(* IEC 61131-3 sources: plc-st-coding-agent/progress/evidence/f14_v10_full_20261113/jobs/custom_minimax-m27 (part 3) *)

(* ---- public-hard-05.raw_candidate_01.st ---- *)
(* CONTRACT_RULES [] *)
FUNCTION_BLOCK ArmController
VAR_INPUT
    ManualMode      : BOOL;
    SingleStepMode  : BOOL;
    SingleCycleMode : BOOL;
    ContinuousMode  : BOOL;
    EmergencyStop   : BOOL;
    Start           : BOOL;
    DownButton      : BOOL;
    UpButton        : BOOL;
    LeftButton      : BOOL;
    RightButton     : BOOL;
    GripButton      : BOOL;
    ReleaseButton   : BOOL;
    DownLimitSwitch : BOOL;
    UpLimitSwitch   : BOOL;
    LeftLimitSwitch : BOOL;
    RightLimitSwitch: BOOL;
    GripLimitSwitch : BOOL;
    ReleaseLimitSwitch: BOOL;
END_VAR
VAR_OUTPUT
    MoveDown        : BOOL;
    MoveUp          : BOOL;
    MoveLeft        : BOOL;
    MoveRight       : BOOL;
    ActivateGrip    : BOOL;
    ActivateRelease : BOOL;
END_VAR
VAR
    tmp_Step : INT := 0;
    tmp_StartPrev : BOOL := FALSE;
    tmp_StartRisingEdge : BOOL;
    tmp_StartReleased : BOOL := FALSE;
    tmp_ActionCompleted : BOOL := FALSE;
END_VAR

(*
ENGINEERING_CONTRACT
====================================================================================================
Output State: Activation | Retention/hold | Explicit reset | Same-scan priority | Units/boundaries
----------------------------------------------------------------------------------------------------
MoveDown:     Manual=button AND NOT limit; Step modes=per step CASE; EmergencyStop→FALSE
MoveUp:       Manual=button AND NOT limit; Step modes=per step CASE; EmergencyStop→FALSE
MoveLeft:     Manual=button AND NOT limit; Step modes=per step CASE; EmergencyStop→FALSE
MoveRight:    Manual=button AND NOT limit; Step modes=per step CASE; EmergencyStop→FALSE
ActivateGrip:     Manual=GripButton; Step modes=per step CASE using GripLimitSwitch; EmergencyStop→FALSE
ActivateRelease:  Manual=ReleaseButton; Step modes=per step CASE using ReleaseLimitSwitch; EmergencyStop→FALSE

Manual Mode (PUB001):
  - Direct button-to-output mapping, held while button pressed and NOT at limit position
  - Grip/Release: held while button pressed (limit switches are feedback only)
  - Priority: Highest; independent of step sequencer state

Single Step Mode (PUB003):
  - Step sequence: Down→Grip→Up→Right→Down→Release→Up→Left→(repeat)
  - Each action requires limit switch confirmation before next Start enables next step
  - Initial arm position: top-left (UpLimitSwitch=1, LeftLimitSwitch=1) [PUB002]
  - Step 0: Wait for Start rising edge, then execute step 1
  - Steps 1-7: Advance when current action completes AND (Start released since last press OR step>0)
  - Step 8: Wait for Start released then pressed again before cycling to step 0

Single Cycle Mode (PUB005):
  - Auto-execute all 8 steps sequentially on single Start press
  - Stops at step 8 (end state) after completing left movement
  - No automatic restart; next Start press required

Continuous Mode (PUB006):
  - Same 8-step sequence as single cycle
  - Automatic restart from step 0 when left movement completes (step→0)
  - Continuous looping until mode change or emergency stop

Emergency Stop (PUB007):
  - Trigger: EmergencyStop=FALSE
  - Effect: All outputs FALSE, step counter reset to 0
  - No automatic resume; requires mode re-activation after E-stop clears

PUB IDs: PUB001, PUB002, PUB003, PUB004, PUB005, PUB006, PUB007, PUB008, PUB009, PUB010, PUB011, PUB012, PUB013, PUB014, PUB015, PUB016, PUB017, PUB018, PUB019, PUB020
====================================================================================================
*)
tmp_StartRisingEdge := Start AND NOT tmp_StartPrev;

MoveDown := FALSE;
MoveUp := FALSE;
MoveLeft := FALSE;
MoveRight := FALSE;
ActivateGrip := FALSE;
ActivateRelease := FALSE;

IF EmergencyStop = FALSE THEN
    MoveDown := FALSE;
    MoveUp := FALSE;
    MoveLeft := FALSE;
    MoveRight := FALSE;
    ActivateGrip := FALSE;
    ActivateRelease := FALSE;
    tmp_Step := 0;
    tmp_StartPrev := Start;
    RETURN;
END_IF;

tmp_StartPrev := Start;

IF ManualMode THEN
    MoveDown := DownButton AND NOT DownLimitSwitch;
    MoveUp := UpButton AND NOT UpLimitSwitch;
    MoveLeft := LeftButton AND NOT LeftLimitSwitch;
    MoveRight := RightButton AND NOT RightLimitSwitch;
    ActivateGrip := GripButton;
    ActivateRelease := ReleaseButton;
ELSIF SingleStepMode THEN
    IF tmp_Step = 0 THEN
        IF tmp_StartRisingEdge THEN
            tmp_Step := 1;
        END_IF;
    ELSIF tmp_Step > 0 THEN
        tmp_ActionCompleted := FALSE;
        CASE tmp_Step OF
            1:
                MoveDown := TRUE;
                IF DownLimitSwitch THEN
                    tmp_ActionCompleted := TRUE;
                END_IF;
            2:
                ActivateGrip := TRUE;
                IF GripLimitSwitch THEN
                    tmp_ActionCompleted := TRUE;
                END_IF;
            3:
                MoveUp := TRUE;
                IF UpLimitSwitch THEN
                    tmp_ActionCompleted := TRUE;
                END_IF;
            4:
                MoveRight := TRUE;
                IF RightLimitSwitch THEN
                    tmp_ActionCompleted := TRUE;
                END_IF;
            5:
                MoveDown := TRUE;
                IF DownLimitSwitch THEN
                    tmp_ActionCompleted := TRUE;
                END_IF;
            6:
                ActivateRelease := TRUE;
                IF ReleaseLimitSwitch THEN
                    tmp_ActionCompleted := TRUE;
                END_IF;
            7:
                MoveUp := TRUE;
                IF UpLimitSwitch THEN
                    tmp_ActionCompleted := TRUE;
                END_IF;
            8:
                MoveLeft := TRUE;
                IF LeftLimitSwitch THEN
                    tmp_ActionCompleted := TRUE;
                END_IF;
        END_CASE;
        IF tmp_ActionCompleted THEN
            tmp_Step := tmp_Step + 1;
            IF tmp_Step > 8 THEN
                tmp_Step := 8;
            END_IF;
            tmp_StartReleased := FALSE;
        END_IF;
        IF NOT Start THEN
            tmp_StartReleased := TRUE;
        END_IF;
        IF tmp_Step = 8 THEN
            IF tmp_StartRisingEdge AND tmp_StartReleased THEN
                tmp_Step := 0;
                tmp_StartReleased := FALSE;
            END_IF;
        ELSIF tmp_StartRisingEdge AND (tmp_StartReleased OR (tmp_Step > 0)) THEN
            tmp_Step := tmp_Step + 1;
            IF tmp_Step > 8 THEN
                tmp_Step := 8;
            END_IF;
            tmp_StartReleased := FALSE;
        END_IF;
    END_IF;
ELSIF SingleCycleMode THEN
    IF tmp_Step = 0 THEN
        IF tmp_StartRisingEdge THEN
            tmp_Step := 1;
        END_IF;
    ELSIF tmp_Step > 0 THEN
        tmp_ActionCompleted := FALSE;
        CASE tmp_Step OF
            1:
                MoveDown := TRUE;
                IF DownLimitSwitch THEN
                    tmp_ActionCompleted := TRUE;
                END_IF;
            2:
                ActivateGrip := TRUE;
                IF GripLimitSwitch THEN
                    tmp_ActionCompleted := TRUE;
                END_IF;
            3:
                MoveUp := TRUE;
                IF UpLimitSwitch THEN
                    tmp_ActionCompleted := TRUE;
                END_IF;
            4:
                MoveRight := TRUE;
                IF RightLimitSwitch THEN
                    tmp_ActionCompleted := TRUE;
                END_IF;
            5:
                MoveDown := TRUE;
                IF DownLimitSwitch THEN
                    tmp_ActionCompleted := TRUE;
                END_IF;
            6:
                ActivateRelease := TRUE;
                IF ReleaseLimitSwitch THEN
                    tmp_ActionCompleted := TRUE;
                END_IF;
            7:
                MoveUp := TRUE;
                IF UpLimitSwitch THEN
                    tmp_ActionCompleted := TRUE;
                END_IF;
            8:
                MoveLeft := TRUE;
                IF LeftLimitSwitch THEN
                    tmp_ActionCompleted := TRUE;
                END_IF;
        END_CASE;
        IF tmp_ActionCompleted THEN
            tmp_Step := tmp_Step + 1;
            IF tmp_Step > 8 THEN
                tmp_Step := 8;
            END_IF;
        END_IF;
    END_IF;
ELSIF ContinuousMode THEN
    IF tmp_Step = 0 THEN
        IF tmp_StartRisingEdge THEN
            tmp_Step := 1;
        END_IF;
    ELSIF tmp_Step > 0 THEN
        tmp_ActionCompleted := FALSE;
        CASE tmp_Step OF
            1:
                MoveDown := TRUE;
                IF DownLimitSwitch THEN
                    tmp_ActionCompleted := TRUE;
                END_IF;
            2:
                ActivateGrip := TRUE;
                IF GripLimitSwitch THEN
                    tmp_ActionCompleted := TRUE;
                END_IF;
            3:
                MoveUp := TRUE;
                IF UpLimitSwitch THEN
                    tmp_ActionCompleted := TRUE;
                END_IF;
            4:
                MoveRight := TRUE;
                IF RightLimitSwitch THEN
                    tmp_ActionCompleted := TRUE;
                END_IF;
            5:
                MoveDown := TRUE;
                IF DownLimitSwitch THEN
                    tmp_ActionCompleted := TRUE;
                END_IF;
            6:
                ActivateRelease := TRUE;
                IF ReleaseLimitSwitch THEN
                    tmp_ActionCompleted := TRUE;
                END_IF;
            7:
                MoveUp := TRUE;
                IF UpLimitSwitch THEN
                    tmp_ActionCompleted := TRUE;
                END_IF;
            8:
                MoveLeft := TRUE;
                IF LeftLimitSwitch THEN
                    tmp_ActionCompleted := TRUE;
                END_IF;
        END_CASE;
        IF tmp_ActionCompleted THEN
            tmp_Step := tmp_Step + 1;
            IF tmp_Step > 8 THEN
                tmp_Step := 0;
            END_IF;
        END_IF;
    END_IF;
END_IF;
END_FUNCTION_BLOCK

(* ---- public-hard-05.raw_candidate_02.st ---- *)
Looking at the checkpoints and test failures, I need to identify the semantics issues:

1. **h05-13 failure**: SingleStepMode, Start=TRUE from previous FALSE state should advance to step 1 (MoveDown=TRUE), but observed is FALSE. This indicates the rising edge `tmp_StartRisingEdge` is not being consumed after use, causing it to persist and advance the step multiple times on the same scan until it passes step 1.

2. The rising edge flag persists across calls when Start remains TRUE, causing `tmp_Step` to skip past 1 before the CASE output assignment executes.

The fix: Clear `tmp_StartRisingEdge` immediately after consuming it at step 0 to ensure single-scan advancement semantics.

(* CONTRACT_RULES [] *)
FUNCTION_BLOCK ArmController
VAR_INPUT
    ManualMode      : BOOL;
    SingleStepMode  : BOOL;
    SingleCycleMode : BOOL;
    ContinuousMode  : BOOL;
    EmergencyStop   : BOOL;
    Start           : BOOL;
    DownButton      : BOOL;
    UpButton        : BOOL;
    LeftButton      : BOOL;
    RightButton     : BOOL;
    GripButton      : BOOL;
    ReleaseButton   : BOOL;
    DownLimitSwitch : BOOL;
    UpLimitSwitch   : BOOL;
    LeftLimitSwitch : BOOL;
    RightLimitSwitch: BOOL;
    GripLimitSwitch : BOOL;
    ReleaseLimitSwitch: BOOL;
END_VAR
VAR_OUTPUT
    MoveDown        : BOOL;
    MoveUp          : BOOL;
    MoveLeft        : BOOL;
    MoveRight       : BOOL;
    ActivateGrip    : BOOL;
    ActivateRelease : BOOL;
END_VAR
VAR
    tmp_Step : INT := 0;
    tmp_StartPrev : BOOL := FALSE;
    tmp_StartRisingEdge : BOOL;
    tmp_StartReleased : BOOL := FALSE;
    tmp_ActionCompleted : BOOL := FALSE;
END_VAR

(*
ENGINEERING_CONTRACT
====================================================================================================
Output State: Activation | Retention/hold | Explicit reset | Same-scan priority | Units/boundaries
----------------------------------------------------------------------------------------------------
MoveDown:     Manual=button AND NOT limit; Step modes=per step CASE; EmergencyStop→FALSE
MoveUp:       Manual=button AND NOT limit; Step modes=per step CASE; EmergencyStop→FALSE
MoveLeft:     Manual=button AND NOT limit; Step modes=per step CASE; EmergencyStop→FALSE
MoveRight:    Manual=button AND NOT limit; Step modes=per step CASE; EmergencyStop→FALSE
ActivateGrip:     Manual=GripButton; Step modes=per step CASE using GripLimitSwitch; EmergencyStop→FALSE
ActivateRelease:  Manual=ReleaseButton; Step modes=per step CASE using ReleaseLimitSwitch; EmergencyStop→FALSE

Manual Mode (PUB001):
  - Direct button-to-output mapping, held while button pressed and NOT at limit position
  - Grip/Release: held while button pressed (limit switches are feedback only)
  - Priority: Highest; independent of step sequencer state

Single Step Mode (PUB003):
  - Step sequence: Down→Grip→Up→Right→Down→Release→Up→Left→(repeat)
  - Each action requires limit switch confirmation before next Start enables next step
  - Initial arm position: top-left (UpLimitSwitch=1, LeftLimitSwitch=1) [PUB002]
  - Step 0: Wait for Start rising edge, then execute step 1
  - Steps 1-7: Advance when current action completes AND (Start released since last press OR step>0)
  - Step 8: Wait for Start released then pressed again before cycling to step 0

Single Cycle Mode (PUB005):
  - Auto-execute all 8 steps sequentially on single Start press
  - Stops at step 8 (end state) after completing left movement
  - No automatic restart; next Start press required

Continuous Mode (PUB006):
  - Same 8-step sequence as single cycle
  - Automatic restart from step 0 when left movement completes (step→0)
  - Continuous looping until mode change or emergency stop

Emergency Stop (PUB007):
  - Trigger: EmergencyStop=FALSE
  - Effect: All outputs FALSE, step counter reset to 0
  - No automatic resume; requires mode re-activation after E-stop clears

PUB IDs: PUB001, PUB002, PUB003, PUB004, PUB005, PUB006, PUB007, PUB008, PUB009, PUB010, PUB011, PUB012, PUB013, PUB014, PUB015, PUB016, PUB017, PUB018, PUB019, PUB020
====================================================================================================
*)
tmp_StartRisingEdge := Start AND NOT tmp_StartPrev;

MoveDown := FALSE;
MoveUp := FALSE;
MoveLeft := FALSE;
MoveRight := FALSE;
ActivateGrip := FALSE;
ActivateRelease := FALSE;

IF EmergencyStop = FALSE THEN
    MoveDown := FALSE;
    MoveUp := FALSE;
    MoveLeft := FALSE;
    MoveRight := FALSE;
    ActivateGrip := FALSE;
    ActivateRelease := FALSE;
    tmp_Step := 0;
    tmp_StartPrev := Start;
    RETURN;
END_IF;

tmp_StartPrev := Start;

IF ManualMode THEN
    MoveDown := DownButton AND NOT DownLimitSwitch;
    MoveUp := UpButton AND NOT UpLimitSwitch;
    MoveLeft := LeftButton AND NOT LeftLimitSwitch;
    MoveRight := RightButton AND NOT RightLimitSwitch;
    ActivateGrip := GripButton;
    ActivateRelease := ReleaseButton;
ELSIF SingleStepMode THEN
    IF tmp_Step = 0 THEN
        IF tmp_StartRisingEdge THEN
            tmp_Step := 1;
            tmp_StartRisingEdge := FALSE;
        END_IF;
    ELSIF tmp_Step > 0 THEN
        tmp_ActionCompleted := FALSE;
        CASE tmp_Step OF
            1:
                MoveDown := TRUE;
                IF DownLimitSwitch THEN
                    tmp_ActionCompleted := TRUE;
                END_IF;
            2:
                ActivateGrip := TRUE;
                IF GripLimitSwitch THEN
                    tmp_ActionCompleted := TRUE;
                END_IF;
            3:
                MoveUp := TRUE;
                IF UpLimitSwitch THEN
                    tmp_ActionCompleted := TRUE;
                END_IF;
            4:
                MoveRight := TRUE;
                IF RightLimitSwitch THEN
                    tmp_ActionCompleted := TRUE;
                END_IF;
            5:
                MoveDown := TRUE;
                IF DownLimitSwitch THEN
                    tmp_ActionCompleted := TRUE;
                END_IF;
            6:
                ActivateRelease := TRUE;
                IF ReleaseLimitSwitch THEN
                    tmp_ActionCompleted := TRUE;
                END_IF;
            7:
                MoveUp := TRUE;
                IF UpLimitSwitch THEN
                    tmp_ActionCompleted := TRUE;
                END_IF;
            8:
                MoveLeft := TRUE;
                IF LeftLimitSwitch THEN
                    tmp_ActionCompleted := TRUE;
                END_IF;
        END_CASE;
        IF tmp_ActionCompleted THEN
            tmp_Step := tmp_Step + 1;
            IF tmp_Step > 8 THEN
                tmp_Step := 8;
            END_IF;
            tmp_StartReleased := FALSE;
        END_IF;
        IF NOT Start THEN
            tmp_StartReleased := TRUE;
        END_IF;
        IF tmp_Step = 8 THEN
            IF tmp_StartRisingEdge AND tmp_StartReleased THEN
                tmp_Step := 0;
                tmp_StartReleased := FALSE;
            END_IF;
        ELSIF tmp_StartRisingEdge AND (tmp_StartReleased OR (tmp_Step > 0)) THEN
            tmp_Step := tmp_Step + 1;
            IF tmp_Step > 8 THEN
                tmp_Step := 8;
            END_IF;
            tmp_StartReleased := FALSE;
        END_IF;
    END_IF;
ELSIF SingleCycleMode THEN
    IF tmp_Step = 0 THEN
        IF tmp_StartRisingEdge THEN
            tmp_Step := 1;
            tmp_StartRisingEdge := FALSE;
        END_IF;
    ELSIF tmp_Step > 0 THEN
        tmp_ActionCompleted := FALSE;
        CASE tmp_Step OF
            1:
                MoveDown := TRUE;
                IF DownLimitSwitch THEN
                    tmp_ActionCompleted := TRUE;
                END_IF;
            2:
                ActivateGrip := TRUE;
                IF GripLimitSwitch THEN
                    tmp_ActionCompleted := TRUE;
                END_IF;
            3:
                MoveUp := TRUE;
                IF UpLimitSwitch THEN
                    tmp_ActionCompleted := TRUE;
                END_IF;
            4:
                MoveRight := TRUE;
                IF RightLimitSwitch THEN
                    tmp_ActionCompleted := TRUE;
                END_IF;
            5:
                MoveDown := TRUE;
                IF DownLimitSwitch THEN
                    tmp_ActionCompleted := TRUE;
                END_IF;
            6:
                ActivateRelease := TRUE;
                IF ReleaseLimitSwitch THEN
                    tmp_ActionCompleted := TRUE;
                END_IF;
            7:
                MoveUp := TRUE;
                IF UpLimitSwitch THEN
                    tmp_ActionCompleted := TRUE;
                END_IF;
            8:
                MoveLeft := TRUE;
                IF LeftLimitSwitch THEN
                    tmp_ActionCompleted := TRUE;
                END_IF;
        END_CASE;
        IF tmp_ActionCompleted THEN
            tmp_Step := tmp_Step + 1;
            IF tmp_Step > 8 THEN
                tmp_Step := 8;
            END_IF;
        END_IF;
    END_IF;
ELSIF ContinuousMode THEN
    IF tmp_Step = 0 THEN
        IF tmp_StartRisingEdge THEN
            tmp_Step := 1;
            tmp_StartRisingEdge := FALSE;
        END_IF;
    ELSIF tmp_Step > 0 THEN
        tmp_ActionCompleted := FALSE;
        CASE tmp_Step OF
            1:
                MoveDown := TRUE;
                IF DownLimitSwitch THEN
                    tmp_ActionCompleted := TRUE;
                END_IF;
            2:
                ActivateGrip := TRUE;
                IF GripLimitSwitch THEN
                    tmp_ActionCompleted := TRUE;
                END_IF;
            3:
                MoveUp := TRUE;
                IF UpLimitSwitch THEN
                    tmp_ActionCompleted := TRUE;
                END_IF;
            4:
                MoveRight := TRUE;
                IF RightLimitSwitch THEN
                    tmp_ActionCompleted := TRUE;
                END_IF;
            5:
                MoveDown := TRUE;
                IF DownLimitSwitch THEN
                    tmp_ActionCompleted := TRUE;
                END_IF;
            6:
                ActivateRelease := TRUE;
                IF ReleaseLimitSwitch THEN
                    tmp_ActionCompleted := TRUE;
                END_IF;
            7:
                MoveUp := TRUE;
                IF UpLimitSwitch THEN
                    tmp_ActionCompleted := TRUE;
                END_IF;
            8:
                MoveLeft := TRUE;
                IF LeftLimitSwitch THEN
                    tmp_ActionCompleted := TRUE;
                END_IF;
        END_CASE;
        IF tmp_ActionCompleted THEN
            tmp_Step := tmp_Step + 1;
            IF tmp_Step > 8 THEN
                tmp_Step := 0;
            END_IF;
        END_IF;
    END_IF;
END_IF;
END_FUNCTION_BLOCK

(* ---- public-hard-06.candidate_01.st ---- *)
(* ENGINEERING_CONTRACT
 * =============================================================================
 * Production Control - 5-Station Automated Line
 * =============================================================================
 * MODES:
 * - Manual (Mode=0): ForwardButton→MotorForward, ReverseButton→MotorReverse
 *   Interlock: MotorForward AND MotorReverse never simultaneous
 *   Activation: Button held; No retention; No explicit reset defined
 *
 * - Automatic (Mode=1): State-machine progression with sensor triggers
 *   States: LOAD→WASH→WEIGH→FIRE→OUTPUT (sequential forward flow)
 *
 * AUTOMATIC STATE TRANSITIONS:
 * - ST_LOAD: SensorFeed → MotorForward (retract, moves to next station)
 *   Reset: Automatic off, manual mode
 *
 * - ST_WASH: SensorWash → MotorStop
 *   Activation: washComplete → MotorForward
 *   Reset: Automatic off, manual mode
 *
 * - ST_WEIGH: SensorWeight → MotorStop
 *   Activation: weightComplete AND qualified(100≤weight≤200) → calc firingTemp, MotorForward
 *   Activation: weightComplete AND NOT qualified → kick latch ON
 *   Reset: Automatic off, manual mode; kick requires external reset (unspecified)
 *
 * - ST_FIRE: SensorFiring → MotorStop
 *   Activation: firingComplete → MotorForward
 *   Reset: Automatic off, manual mode
 *
 * - ST_OUTPUT: SensorOutput → MotorStop, CompletionLight:=SensorOutput
 *   Retention: CompletionLight held ON while SensorOutput=TRUE; OFF when FALSE
 *   Reset: Automatic off, manual mode (light follows sensor)
 *
 * FIRING TEMP CALCULATION:
 * - Linear: weight 100→200 maps to temp 500→550
 * - Formula: firingTemp = 500.0 + (weight - 100.0) * 0.5
 * - Only calculated once per qualified product (on weightComplete)
 * - Retained until next qualified product (unspecified reset)
 *
 * UNITS/BOUNDARIES:
 * - Weight: REAL, qualified range [100.0, 200.0] inclusive
 * - Temp: REAL, output range [500.0, 550.0] inclusive
 * - All sensors: BOOL, edge-triggered detection (sensor TRUE = product arrived)
 * =============================================================================
 *)

(* CONTRACT_RULES [{"kind":"hold_until_reset","output":"kick","set_input":"weightComplete","reset_input":null}] *)

FUNCTION_BLOCK ProductionControl
VAR_INPUT
    Mode            : BOOL;  (* 0=manual, 1=automatic *)
    ForwardButton   : BOOL;
    ReverseButton   : BOOL;
    SensorFeed      : BOOL;
    SensorWash      : BOOL;
    SensorWeight    : BOOL;
    SensorFiring    : BOOL;
    SensorOutput    : BOOL;
    washComplete    : BOOL;
    weightComplete  : BOOL;
    weight          : REAL;
    firingComplete  : BOOL;
END_VAR

VAR_OUTPUT
    MotorForward    : BOOL;
    MotorReverse    : BOOL;
    kick            : BOOL;
    CompletionLight : BOOL;
    firingTemp      : REAL;
END_VAR

VAR
    state           : INT;   (* 0=LOAD, 1=WASH, 2=WEIGH, 3=FIRE, 4=OUTPUT *)
    prevWashComplete    : BOOL;
    prevWeightComplete  : BOOL;
    prevFiringComplete  : BOOL;
    tmp_Qualified       : BOOL;
    tmp_TempCalc        : REAL;
END_VAR

(* State constants *)
CONST
    ST_LOAD   := 0;
    ST_WASH   := 1;
    ST_WEIGH  := 2;
    ST_FIRE   := 3;
    ST_OUTPUT := 4;
END_CONST

(* Initialize outputs to safe state *)
MotorForward    := FALSE;
MotorReverse    := FALSE;
kick            := kick;        (* Preserve retained state *)
CompletionLight := FALSE;
firingTemp      := firingTemp;  (* Preserve retained state *)

IF Mode = FALSE THEN
    (* ======================================================================= *)
    (* MANUAL MODE                                                             *)
    (* PUB001, PUB002, PUB003                                                  *)
    (* ======================================================================= *)
    (* Interlock: forward and reverse cannot be simultaneous *)
    IF ForwardButton AND NOT ReverseButton THEN
        MotorForward := TRUE;
        MotorReverse := FALSE;
    ELSIF ReverseButton AND NOT ForwardButton THEN
        MotorForward := FALSE;
        MotorReverse := TRUE;
    ELSE
        MotorForward := FALSE;
        MotorReverse := FALSE;
    END_IF;

    (* Reset state machine when entering manual mode *)
    state := ST_LOAD;

ELSIF Mode = TRUE THEN
    (* ======================================================================= *)
    (* AUTOMATIC MODE                                                          *)
    (* PUB004, PUB005, PUB006, PUB007, PUB008, PUB009, PUB010, PUB011, PUB012   *)
    (* ======================================================================= *)
    MotorReverse := FALSE;  (* Only forward in automatic mode *)

    (* Edge detection for completion signals *)
    IF washComplete AND NOT prevWashComplete THEN
        (* Rising edge on washComplete *)
        MotorForward := TRUE;
    END_IF;
    prevWashComplete := washComplete;

    IF firingComplete AND NOT prevFiringComplete THEN
        (* Rising edge on firingComplete *)
        MotorForward := TRUE;
    END_IF;
    prevFiringComplete := firingComplete;

    (* State machine based on current station detection *)
    IF SensorOutput THEN
        (* ================================================================= *)
        (* STATION 5: OUTPUT (Finished Product)                              *)
        (* PUB012                                                              *)
        (* Motor stops, CompletionLight follows sensor                       *)
        (* ================================================================= *)
        state := ST_OUTPUT;
        MotorForward := FALSE;
        CompletionLight := SensorOutput;  (* ON when product present *)

    ELSIF SensorFiring THEN
        (* ================================================================= *)
        (* STATION 4: FIRING                                                 *)
        (* PUB010, PUB011                                                     *)
        (* Motor stops; wait for firingComplete → forward                    *)
        (* ================================================================= *)
        state := ST_FIRE;
        MotorForward := FALSE;
        CompletionLight := FALSE;
        (* MotorForward set on rising edge of firingComplete above *)

    ELSIF SensorWeight THEN
        (* ================================================================= *)
        (* STATION 3: WEIGHING                                                *)
        (* PUB006, PUB007, PUB008, PUB009                                     *)
        (* Motor stops; weightComplete triggers qualification check           *)
        (* ================================================================= *)
        state := ST_WEIGH;
        MotorForward := FALSE;
        CompletionLight := FALSE;

        (* Rising edge detection for weightComplete *)
        IF weightComplete AND NOT prevWeightComplete THEN
            prevWeightComplete := weightComplete;

            (* Qualification check: 100 <= weight <= 200 *)
            IF weight >= 100.0 AND weight <= 200.0 THEN
                (* Qualified: calculate firing temperature *)
                (* Linear interpolation: weight[100,200] -> temp[500,550] *)
                tmp_TempCalc := 500.0 + (weight - 100.0) * 0.5;
                firingTemp := tmp_TempCalc;
                kick := FALSE;
                MotorForward := TRUE;
            ELSE
                (* Unqualified: reject *)
                kick := TRUE;
                MotorForward := FALSE;
            END_IF;
        ELSE
            prevWeightComplete := weightComplete;
        END_IF;

    ELSIF SensorWash THEN
        (* ================================================================= *)
        (* STATION 2: CLEANING                                                *)
        (* PUB004, PUB005                                                     *)
        (* Motor stops; washComplete triggers forward                        *)
        (* ================================================================= *)
        state := ST_WASH;
        MotorForward := FALSE;
        CompletionLight := FALSE;
        kick := FALSE;  (* Reset kick on new product entering wash *)

    ELSIF SensorFeed THEN
        (* ================================================================= *)
        (* STATION 1: MATERIAL LOADING                                        *)
        (* PUB004                                                              *)
        (* SensorFeed detected → start motor forward                         *)
        (* ================================================================= *)
        state := ST_LOAD;
        MotorForward := TRUE;
        CompletionLight := FALSE;
        kick := FALSE;  (* Reset kick on new product *)

    ELSE
        (* No sensor active - product in transit or line empty *)
        (* Maintain current MotorForward state from completion signals *)
        (* MotorForward already set by rising edges above *)
        CompletionLight := FALSE;
    END_IF;

END_IF;

END_FUNCTION_BLOCK

(* ---- public-hard-06.candidate_02.st ---- *)
(* ENGINEERING_CONTRACT
 * =============================================================================
 * Production Control - 5-Station Automated Line
 * =============================================================================
 * MODES:
 * - Manual (Mode=0): ForwardButton→MotorForward, ReverseButton→MotorReverse
 *   Interlock: MotorForward AND MotorReverse never simultaneous
 *   Activation: Button held; No retention; No explicit reset defined
 *
 * - Automatic (Mode=1): State-machine progression with sensor triggers
 *   States: LOAD→WASH→WEIGH→FIRE→OUTPUT (sequential forward flow)
 *
 * AUTOMATIC STATE TRANSITIONS:
 * - ST_LOAD: SensorFeed → MotorForward (retract, moves to next station)
 *   Reset: Automatic off, manual mode
 *
 * - ST_WASH: SensorWash → MotorStop
 *   Activation: washComplete → MotorForward
 *   Reset: Automatic off, manual mode
 *
 * - ST_WEIGH: SensorWeight → MotorStop
 *   Activation: weightComplete AND qualified(100≤weight≤200) → calc firingTemp, MotorForward
 *   Activation: weightComplete AND NOT qualified → kick latch ON
 *   Reset: Automatic off, manual mode; kick requires external reset (unspecified)
 *
 * - ST_FIRE: SensorFiring → MotorStop
 *   Activation: firingComplete → MotorForward
 *   Reset: Automatic off, manual mode
 *
 * - ST_OUTPUT: SensorOutput → MotorStop, CompletionLight:=SensorOutput
 *   Retention: CompletionLight held ON while SensorOutput=TRUE; OFF when FALSE
 *   Reset: Automatic off, manual mode (light follows sensor)
 *
 * FIRING TEMP CALCULATION:
 * - Linear: weight 100→200 maps to temp 500→550
 * - Formula: firingTemp = 500.0 + (weight - 100.0) * 0.5
 * - Only calculated once per qualified product (on weightComplete)
 * - Retained until next qualified product (unspecified reset)
 *
 * UNITS/BOUNDARIES:
 * - Weight: REAL, qualified range [100.0, 200.0] inclusive
 * - Temp: REAL, output range [500.0, 550.0] inclusive
 * - All sensors: BOOL, edge-triggered detection (sensor TRUE = product arrived)
 * =============================================================================
 *)

(* CONTRACT_RULES [{"kind":"hold_until_reset","output":"kick","set_input":"weightComplete","reset_input":null}] *)

TYPE StationState :
(
    ST_LOAD   := 0,
    ST_WASH   := 1,
    ST_WEIGH  := 2,
    ST_FIRE   := 3,
    ST_OUTPUT := 4
);
END_TYPE;

FUNCTION_BLOCK ProductionControl
VAR_INPUT
    Mode            : BOOL;  (* 0=manual, 1=automatic *)
    ForwardButton   : BOOL;
    ReverseButton   : BOOL;
    SensorFeed      : BOOL;
    SensorWash      : BOOL;
    SensorWeight    : BOOL;
    SensorFiring    : BOOL;
    SensorOutput    : BOOL;
    washComplete    : BOOL;
    weightComplete  : BOOL;
    weight          : REAL;
    firingComplete  : BOOL;
END_VAR

VAR_OUTPUT
    MotorForward    : BOOL;
    MotorReverse    : BOOL;
    kick            : BOOL;
    CompletionLight : BOOL;
    firingTemp      : REAL;
END_VAR

VAR
    state               : StationState;
    prevWashComplete    : BOOL;
    prevWeightComplete  : BOOL;
    prevFiringComplete  : BOOL;
    tmp_Qualified       : BOOL;
    tmp_TempCalc        : REAL;
END_VAR

(* Initialize outputs to safe state *)
MotorForward    := FALSE;
MotorReverse    := FALSE;
kick            := kick;        (* Preserve retained state *)
CompletionLight := FALSE;
firingTemp      := firingTemp;  (* Preserve retained state *)

IF Mode = FALSE THEN
    (* ======================================================================= *)
    (* MANUAL MODE                                                             *)
    (* PUB001, PUB002, PUB003                                                  *)
    (* ======================================================================= *)
    (* Interlock: forward and reverse cannot be simultaneous *)
    IF ForwardButton AND NOT ReverseButton THEN
        MotorForward := TRUE;
        MotorReverse := FALSE;
    ELSIF ReverseButton AND NOT ForwardButton THEN
        MotorForward := FALSE;
        MotorReverse := TRUE;
    ELSE
        MotorForward := FALSE;
        MotorReverse := FALSE;
    END_IF;

    (* Reset state machine when entering manual mode *)
    state := ST_LOAD;

ELSIF Mode = TRUE THEN
    (* ======================================================================= *)
    (* AUTOMATIC MODE                                                          *)
    (* PUB004, PUB005, PUB006, PUB007, PUB008, PUB009, PUB010, PUB011, PUB012   *)
    (* ======================================================================= *)
    MotorReverse := FALSE;  (* Only forward in automatic mode *)

    (* Edge detection for completion signals *)
    IF washComplete AND NOT prevWashComplete THEN
        (* Rising edge on washComplete *)
        MotorForward := TRUE;
    END_IF;
    prevWashComplete := washComplete;

    IF firingComplete AND NOT prevFiringComplete THEN
        (* Rising edge on firingComplete *)
        MotorForward := TRUE;
    END_IF;
    prevFiringComplete := firingComplete;

    (* State machine based on current station detection *)
    IF SensorOutput THEN
        (* ================================================================= *)
        (* STATION 5: OUTPUT (Finished Product)                              *)
        (* PUB012                                                              *)
        (* Motor stops, CompletionLight follows sensor                       *)
        (* ================================================================= *)
        state := ST_OUTPUT;
        MotorForward := FALSE;
        CompletionLight := SensorOutput;  (* ON when product present *)

    ELSIF SensorFiring THEN
        (* ================================================================= *)
        (* STATION 4: FIRING                                                 *)
        (* PUB010, PUB011                                                     *)
        (* Motor stops; wait for firingComplete → forward                    *)
        (* ================================================================= *)
        state := ST_FIRE;
        MotorForward := FALSE;
        CompletionLight := FALSE;
        (* MotorForward set on rising edge of firingComplete above *)

    ELSIF SensorWeight THEN
        (* ================================================================= *)
        (* STATION 3: WEIGHING                                                *)
        (* PUB006, PUB007, PUB008, PUB009                                     *)
        (* Motor stops; weightComplete triggers qualification check           *)
        (* ================================================================= *)
        state := ST_WEIGH;
        MotorForward := FALSE;
        CompletionLight := FALSE;

        (* Rising edge detection for weightComplete *)
        IF weightComplete AND NOT prevWeightComplete THEN
            prevWeightComplete := weightComplete;

            (* Qualification check: 100 <= weight <= 200 *)
            IF weight >= 100.0 AND weight <= 200.0 THEN
                (* Qualified: calculate firing temperature *)
                (* Linear interpolation: weight[100,200] -> temp[500,550] *)
                tmp_TempCalc := 500.0 + (weight - 100.0) * 0.5;
                firingTemp := tmp_TempCalc;
                kick := FALSE;
                MotorForward := TRUE;
            ELSE
                (* Unqualified: reject *)
                kick := TRUE;
                MotorForward := FALSE;
            END_IF;
        ELSE
            prevWeightComplete := weightComplete;
        END_IF;

    ELSIF SensorWash THEN
        (* ================================================================= *)
        (* STATION 2: CLEANING                                                *)
        (* PUB004, PUB005                                                     *)
        (* Motor stops; washComplete triggers forward                        *)
        (* ================================================================= *)
        state := ST_WASH;
        MotorForward := FALSE;
        CompletionLight := FALSE;
        kick := FALSE;  (* Reset kick on new product entering wash *)

    ELSIF SensorFeed THEN
        (* ================================================================= *)
        (* STATION 1: MATERIAL LOADING                                        *)
        (* PUB004                                                              *)
        (* SensorFeed detected → start motor forward                         *)
        (* ================================================================= *)
        state := ST_LOAD;
        MotorForward := TRUE;
        CompletionLight := FALSE;
        kick := FALSE;  (* Reset kick on new product *)

    ELSE
        (* No sensor active - product in transit or line empty *)
        (* Maintain current MotorForward state from completion signals *)
        (* MotorForward already set by rising edges above *)
        CompletionLight := FALSE;
    END_IF;

END_IF;

END_FUNCTION_BLOCK

(* ---- public-hard-06.candidate_03.st ---- *)
(* ENGINEERING_CONTRACT
 * =============================================================================
 * Production Control - 5-Station Automated Line
 * =============================================================================
 * MODES:
 * - Manual (Mode=0): ForwardButton→MotorForward, ReverseButton→MotorReverse
 *   Interlock: MotorForward AND MotorReverse never simultaneous
 *   Activation: Button held; No retention; No explicit reset defined
 *
 * - Automatic (Mode=1): State-machine progression with sensor triggers
 *   States: LOAD→WASH→WEIGH→FIRE→OUTPUT (sequential forward flow)
 *
 * AUTOMATIC STATE TRANSITIONS:
 * - ST_LOAD: SensorFeed → MotorForward (retract, moves to next station)
 *   Reset: Automatic off, manual mode
 *
 * - ST_WASH: SensorWash → MotorStop
 *   Activation: washComplete → MotorForward
 *   Reset: Automatic off, manual mode
 *
 * - ST_WEIGH: SensorWeight → MotorStop
 *   Activation: weightComplete AND qualified(100≤weight≤200) → calc firingTemp, MotorForward
 *   Activation: weightComplete AND NOT qualified → kick latch ON
 *   Reset: Automatic off, manual mode; kick requires external reset (unspecified)
 *
 * - ST_FIRE: SensorFiring → MotorStop
 *   Activation: firingComplete → MotorForward
 *   Reset: Automatic off, manual mode
 *
 * - ST_OUTPUT: SensorOutput → MotorStop, CompletionLight:=SensorOutput
 *   Retention: CompletionLight held ON while SensorOutput=TRUE; OFF when FALSE
 *   Reset: Automatic off, manual mode (light follows sensor)
 *
 * FIRING TEMP CALCULATION:
 * - Linear: weight 100→200 maps to temp 500→550
 * - Formula: firingTemp = 500.0 + (weight - 100.0) * 0.5
 * - Same-scan calculation when SensorWeight AND weightComplete both TRUE
 * - Retained until next qualified product (unspecified reset)
 *
 * UNITS/BOUNDARIES:
 * - Weight: REAL, qualified range [100.0, 200.0] inclusive
 * - Temp: REAL, output range [500.0, 550.0] inclusive
 * - All sensors: BOOL, level-triggered detection (sensor TRUE = product present)
 * =============================================================================
 *)

(* CONTRACT_RULES [] *)

TYPE StationState :
(
    ST_LOAD   := 0,
    ST_WASH   := 1,
    ST_WEIGH  := 2,
    ST_FIRE   := 3,
    ST_OUTPUT := 4
);
END_TYPE;

FUNCTION_BLOCK ProductionControl
VAR_INPUT
    Mode            : BOOL;  (* 0=manual, 1=automatic *)
    ForwardButton   : BOOL;
    ReverseButton   : BOOL;
    SensorFeed      : BOOL;
    SensorWash      : BOOL;
    SensorWeight    : BOOL;
    SensorFiring    : BOOL;
    SensorOutput    : BOOL;
    washComplete    : BOOL;
    weightComplete  : BOOL;
    weight          : REAL;
    firingComplete  : BOOL;
END_VAR

VAR_OUTPUT
    MotorForward    : BOOL;
    MotorReverse    : BOOL;
    kick             : BOOL;
    CompletionLight : BOOL;
    firingTemp      : REAL;
END_VAR

VAR
    state              : StationState;
    prevWashComplete   : BOOL;
    prevFiringComplete : BOOL;
END_VAR

(* Initialize outputs to safe state *)
MotorForward    := FALSE;
MotorReverse    := FALSE;
kick            := kick;        (* Preserve retained state *)
CompletionLight := FALSE;
firingTemp      := firingTemp;  (* Preserve retained state *)

IF Mode = FALSE THEN
    (* ======================================================================= *)
    (* MANUAL MODE                                                             *)
    (* PUB001, PUB002, PUB003                                                  *)
    (* ======================================================================= *)
    (* Interlock: forward and reverse cannot be simultaneous *)
    IF ForwardButton AND NOT ReverseButton THEN
        MotorForward := TRUE;
        MotorReverse := FALSE;
    ELSIF ReverseButton AND NOT ForwardButton THEN
        MotorForward := FALSE;
        MotorReverse := TRUE;
    ELSE
        MotorForward := FALSE;
        MotorReverse := FALSE;
    END_IF;

    (* Reset state machine when entering manual mode *)
    state := ST_LOAD;

ELSIF Mode = TRUE THEN
    (* ======================================================================= *)
    (* AUTOMATIC MODE                                                          *)
    (* PUB004, PUB005, PUB006, PUB007, PUB008, PUB009, PUB010, PUB011, PUB012   *)
    (* ======================================================================= *)
    MotorReverse := FALSE;  (* Only forward in automatic mode *)

    (* Edge detection for washComplete - rising edge triggers forward *)
    IF washComplete AND NOT prevWashComplete THEN
        MotorForward := TRUE;
    END_IF;
    prevWashComplete := washComplete;

    (* Edge detection for firingComplete - rising edge triggers forward *)
    IF firingComplete AND NOT prevFiringComplete THEN
        MotorForward := TRUE;
    END_IF;
    prevFiringComplete := firingComplete;

    (* State machine based on current station detection *)
    IF SensorOutput THEN
        (* ================================================================= *)
        (* STATION 5: OUTPUT (Finished Product)                              *)
        (* PUB012                                                              *)
        (* Motor stops, CompletionLight follows sensor                       *)
        (* ================================================================= *)
        state := ST_OUTPUT;
        MotorForward := FALSE;
        CompletionLight := SensorOutput;  (* ON when product present *)

    ELSIF SensorFiring THEN
        (* ================================================================= *)
        (* STATION 4: FIRING                                                 *)
        (* PUB010, PUB011                                                     *)
        (* Motor stops; wait for firingComplete → forward                    *)
        (* ================================================================= *)
        state := ST_FIRE;
        MotorForward := FALSE;
        CompletionLight := FALSE;
        (* MotorForward set on rising edge of firingComplete above *)

    ELSIF SensorWeight THEN
        (* ================================================================= *)
        (* STATION 3: WEIGHING                                                *)
        (* PUB006, PUB007, PUB008, PUB009                                     *)
        (* Motor stops; weightComplete triggers qualification check           *)
        (* ================================================================= *)
        state := ST_WEIGH;
        MotorForward := FALSE;
        CompletionLight := FALSE;

        (* Immediate calculation when weightComplete signal is received *)
        (* No edge delay - weightComplete is a one-shot from external process *)
        IF weightComplete THEN
            (* Qualification check: 100 <= weight <= 200 *)
            IF weight >= 100.0 AND weight <= 200.0 THEN
                (* Qualified: calculate firing temperature *)
                (* Linear interpolation: weight[100,200] -> temp[500,550] *)
                firingTemp := 500.0 + (weight - 100.0) * 0.5;
                kick := FALSE;
                MotorForward := TRUE;
            ELSE
                (* Unqualified: reject *)
                kick := TRUE;
                MotorForward := FALSE;
            END_IF;
        END_IF;

    ELSIF SensorWash THEN
        (* ================================================================= *)
        (* STATION 2: CLEANING                                                *)
        (* PUB004, PUB005                                                     *)
        (* Motor stops; washComplete triggers forward                        *)
        (* ================================================================= *)
        state := ST_WASH;
        MotorForward := FALSE;
        CompletionLight := FALSE;
        kick := FALSE;  (* Reset kick on new product entering wash *)

    ELSIF SensorFeed THEN
        (* ================================================================= *)
        (* STATION 1: MATERIAL LOADING                                        *)
        (* PUB004                                                              *)
        (* SensorFeed detected → start motor forward                         *)
        (* ================================================================= *)
        state := ST_LOAD;
        MotorForward := TRUE;
        CompletionLight := FALSE;
        kick := FALSE;  (* Reset kick on new product *)

    ELSE
        (* No sensor active - product in transit or line empty *)
        (* Maintain current MotorForward state from completion signals *)
        (* MotorForward already set by rising edges above *)
        CompletionLight := FALSE;
    END_IF;

END_IF;

END_FUNCTION_BLOCK

(* ---- public-hard-06.candidate_04.st ---- *)
(* ENGINEERING_CONTRACT
 * Production Control - 5-Station Line
 * =============================================================================
 * MODES:
 * - Manual (Mode=0): ForwardButton→MotorForward, ReverseButton→MotorReverse
 *   Interlock: MotorForward AND MotorReverse never simultaneous
 *   Activation: Button held; No retention; No explicit reset defined
 *
 * - Automatic (Mode=1): State-machine progression with sensor triggers
 *   States: LOAD→WASH→WEIGH→FIRE→OUTPUT (sequential forward flow)
 *
 * AUTOMATIC STATE TRANSITIONS:
 * - ST_LOAD: SensorFeed → MotorForward (moves to cleaning station)
 * - ST_WASH: SensorWash → MotorStop; washComplete rising edge → MotorForward
 * - ST_WEIGH: SensorWeight → MotorStop; weightComplete rising edge:
 *   • weight in [100,200] → calc firingTemp (500+0.5*(w-100)), MotorForward
 *   • weight outside range → kick:=TRUE
 * - ST_FIRE: SensorFiring → MotorStop; firingComplete rising edge → MotorForward
 * - ST_OUTPUT: SensorOutput → MotorStop, CompletionLight:=SensorOutput
 *
 * UNITS/BOUNDARIES: Weight REAL in [100,200], Temp REAL in [500,550]
 * =============================================================================
 *)

(* CONTRACT_RULES [{"kind":"hold_until_reset","output":"kick","set_input":"weightComplete","reset_input":null}] *)

TYPE StationState :
(
    ST_LOAD   := 0,
    ST_WASH   := 1,
    ST_WEIGH  := 2,
    ST_FIRE   := 3,
    ST_OUTPUT := 4
);
END_TYPE;

FUNCTION_BLOCK ProductionControl
VAR_INPUT
    Mode            : BOOL;
    ForwardButton   : BOOL;
    ReverseButton   : BOOL;
    SensorFeed      : BOOL;
    SensorWash      : BOOL;
    SensorWeight    : BOOL;
    SensorFiring    : BOOL;
    SensorOutput    : BOOL;
    washComplete    : BOOL;
    weightComplete  : BOOL;
    weight          : REAL;
    firingComplete  : BOOL;
END_VAR

VAR_OUTPUT
    MotorForward    : BOOL;
    MotorReverse    : BOOL;
    kick            : BOOL;
    CompletionLight : BOOL;
    firingTemp      : REAL;
END_VAR

VAR
    state               : StationState;
    prevWashComplete    : BOOL;
    prevWeightComplete  : BOOL;
    prevFiringComplete  : BOOL;
    tmp_MotorForwardCmd : BOOL;
END_VAR

(* Rising edge detection - evaluate BEFORE any state transitions *)
VAR
    washCompleteRising   : BOOL;
    weightCompleteRising : BOOL;
    firingCompleteRising : BOOL;
END_VAR

washCompleteRising   := washComplete   AND NOT prevWashComplete;
weightCompleteRising := weightComplete AND NOT prevWeightComplete;
firingCompleteRising := firingComplete AND NOT prevFiringComplete;

(* Update previous states AFTER edge detection *)
prevWashComplete   := washComplete;
prevWeightComplete := weightComplete;
prevFiringComplete := firingComplete;

(* Default outputs - safety state *)
MotorForward    := FALSE;
MotorReverse    := FALSE;
CompletionLight := FALSE;

IF Mode = FALSE THEN
    (* ======================================================================= *)
    (* MANUAL MODE - PUB001, PUB002, PUB003                                    *)
    (* ======================================================================= *)
    IF ForwardButton AND NOT ReverseButton THEN
        MotorForward := TRUE;
        MotorReverse := FALSE;
    ELSIF ReverseButton AND NOT ForwardButton THEN
        MotorForward := FALSE;
        MotorReverse := TRUE;
    ELSE
        MotorForward := FALSE;
        MotorReverse := FALSE;
    END_IF;

    state := ST_LOAD;

ELSE
    (* ======================================================================= *)
    (* AUTOMATIC MODE - PUB004-PUB012                                           *)
    (* ======================================================================= *)
    MotorReverse := FALSE;

    (* Completion edges set motor forward command - takes priority *)
    IF washCompleteRising THEN
        tmp_MotorForwardCmd := TRUE;
    ELSIF firingCompleteRising THEN
        tmp_MotorForwardCmd := TRUE;
    ELSE
        tmp_MotorForwardCmd := FALSE;
    END_IF;

    (* Kick latch: activated on weightComplete rising edge per contract *)
    IF weightCompleteRising THEN
        IF weight >= 100.0 AND weight <= 200.0 THEN
            kick := FALSE;
        ELSE
            kick := TRUE;
        END_IF;
    END_IF;

    (* Firing temp: calculated on weightComplete rising edge for qualified weight *)
    IF weightCompleteRising THEN
        IF weight >= 100.0 AND weight <= 200.0 THEN
            firingTemp := 500.0 + (weight - 100.0) * 0.5;
        END_IF;
    END_IF;

    (* State machine based on sensor detection *)
    IF SensorOutput THEN
        state := ST_OUTPUT;
        tmp_MotorForwardCmd := FALSE;
        CompletionLight := TRUE;

    ELSIF SensorFiring THEN
        state := ST_FIRE;
        (* Only clear if no completion edge overrode *)
        IF NOT firingCompleteRising THEN
            tmp_MotorForwardCmd := FALSE;
        END_IF;
        CompletionLight := FALSE;

    ELSIF SensorWeight THEN
        state := ST_WEIGH;
        IF NOT weightCompleteRising THEN
            tmp_MotorForwardCmd := FALSE;
        END_IF;
        CompletionLight := FALSE;

    ELSIF SensorWash THEN
        state := ST_WASH;
        IF NOT washCompleteRising THEN
            tmp_MotorForwardCmd := FALSE;
        END_IF;
        CompletionLight := FALSE;

    ELSIF SensorFeed THEN
        state := ST_LOAD;
        tmp_MotorForwardCmd := TRUE;
        CompletionLight := FALSE;
        kick := FALSE;

    ELSE
        (* No sensor active - product in transit *)
        CompletionLight := FALSE;
    END_IF;

END_IF;

(* Apply accumulated motor forward command *)
MotorForward := tmp_MotorForwardCmd;

END_FUNCTION_BLOCK

(* ---- public-hard-06.raw_candidate_01.st ---- *)
(* ENGINEERING_CONTRACT
 * =============================================================================
 * Production Control - 5-Station Automated Line
 * =============================================================================
 * MODES:
 * - Manual (Mode=0): ForwardButton→MotorForward, ReverseButton→MotorReverse
 *   Interlock: MotorForward AND MotorReverse never simultaneous
 *   Activation: Button held; No retention; No explicit reset defined
 *
 * - Automatic (Mode=1): State-machine progression with sensor triggers
 *   States: LOAD→WASH→WEIGH→FIRE→OUTPUT (sequential forward flow)
 *
 * AUTOMATIC STATE TRANSITIONS:
 * - ST_LOAD: SensorFeed → MotorForward (retract, moves to next station)
 *   Reset: Automatic off, manual mode
 *
 * - ST_WASH: SensorWash → MotorStop
 *   Activation: washComplete → MotorForward
 *   Reset: Automatic off, manual mode
 *
 * - ST_WEIGH: SensorWeight → MotorStop
 *   Activation: weightComplete AND qualified(100≤weight≤200) → calc firingTemp, MotorForward
 *   Activation: weightComplete AND NOT qualified → kick latch ON
 *   Reset: Automatic off, manual mode; kick requires external reset (unspecified)
 *
 * - ST_FIRE: SensorFiring → MotorStop
 *   Activation: firingComplete → MotorForward
 *   Reset: Automatic off, manual mode
 *
 * - ST_OUTPUT: SensorOutput → MotorStop, CompletionLight:=SensorOutput
 *   Retention: CompletionLight held ON while SensorOutput=TRUE; OFF when FALSE
 *   Reset: Automatic off, manual mode (light follows sensor)
 *
 * FIRING TEMP CALCULATION:
 * - Linear: weight 100→200 maps to temp 500→550
 * - Formula: firingTemp = 500.0 + (weight - 100.0) * 0.5
 * - Only calculated once per qualified product (on weightComplete)
 * - Retained until next qualified product (unspecified reset)
 *
 * UNITS/BOUNDARIES:
 * - Weight: REAL, qualified range [100.0, 200.0] inclusive
 * - Temp: REAL, output range [500.0, 550.0] inclusive
 * - All sensors: BOOL, edge-triggered detection (sensor TRUE = product arrived)
 * =============================================================================
 *)

(* CONTRACT_RULES [{"kind":"hold_until_reset","output":"kick","set_input":"weightComplete","reset_input":null}] *)

FUNCTION_BLOCK ProductionControl
VAR_INPUT
    Mode            : BOOL;  (* 0=manual, 1=automatic *)
    ForwardButton   : BOOL;
    ReverseButton   : BOOL;
    SensorFeed      : BOOL;
    SensorWash      : BOOL;
    SensorWeight    : BOOL;
    SensorFiring    : BOOL;
    SensorOutput    : BOOL;
    washComplete    : BOOL;
    weightComplete  : BOOL;
    weight          : REAL;
    firingComplete  : BOOL;
END_VAR

VAR_OUTPUT
    MotorForward    : BOOL;
    MotorReverse    : BOOL;
    kick            : BOOL;
    CompletionLight : BOOL;
    firingTemp      : REAL;
END_VAR

VAR
    state           : INT;   (* 0=LOAD, 1=WASH, 2=WEIGH, 3=FIRE, 4=OUTPUT *)
    prevWashComplete    : BOOL;
    prevWeightComplete  : BOOL;
    prevFiringComplete  : BOOL;
    tmp_Qualified       : BOOL;
    tmp_TempCalc        : REAL;
END_VAR

(* State constants *)
CONST
    ST_LOAD   := 0;
    ST_WASH   := 1;
    ST_WEIGH  := 2;
    ST_FIRE   := 3;
    ST_OUTPUT := 4;
END_CONST

(* Initialize outputs to safe state *)
MotorForward    := FALSE;
MotorReverse    := FALSE;
kick            := kick;        (* Preserve retained state *)
CompletionLight := FALSE;
firingTemp      := firingTemp;  (* Preserve retained state *)

IF Mode = FALSE THEN
    (* ======================================================================= *)
    (* MANUAL MODE                                                             *)
    (* PUB001, PUB002, PUB003                                                  *)
    (* ======================================================================= *)
    (* Interlock: forward and reverse cannot be simultaneous *)
    IF ForwardButton AND NOT ReverseButton THEN
        MotorForward := TRUE;
        MotorReverse := FALSE;
    ELSIF ReverseButton AND NOT ForwardButton THEN
        MotorForward := FALSE;
        MotorReverse := TRUE;
    ELSE
        MotorForward := FALSE;
        MotorReverse := FALSE;
    END_IF;

    (* Reset state machine when entering manual mode *)
    state := ST_LOAD;

ELSIF Mode = TRUE THEN
    (* ======================================================================= *)
    (* AUTOMATIC MODE                                                          *)
    (* PUB004, PUB005, PUB006, PUB007, PUB008, PUB009, PUB010, PUB011, PUB012   *)
    (* ======================================================================= *)
    MotorReverse := FALSE;  (* Only forward in automatic mode *)

    (* Edge detection for completion signals *)
    IF washComplete AND NOT prevWashComplete THEN
        (* Rising edge on washComplete *)
        MotorForward := TRUE;
    END_IF;
    prevWashComplete := washComplete;

    IF firingComplete AND NOT prevFiringComplete THEN
        (* Rising edge on firingComplete *)
        MotorForward := TRUE;
    END_IF;
    prevFiringComplete := firingComplete;

    (* State machine based on current station detection *)
    IF SensorOutput THEN
        (* ================================================================= *)
        (* STATION 5: OUTPUT (Finished Product)                              *)
        (* PUB012                                                              *)
        (* Motor stops, CompletionLight follows sensor                       *)
        (* ================================================================= *)
        state := ST_OUTPUT;
        MotorForward := FALSE;
        CompletionLight := SensorOutput;  (* ON when product present *)

    ELSIF SensorFiring THEN
        (* ================================================================= *)
        (* STATION 4: FIRING                                                 *)
        (* PUB010, PUB011                                                     *)
        (* Motor stops; wait for firingComplete → forward                    *)
        (* ================================================================= *)
        state := ST_FIRE;
        MotorForward := FALSE;
        CompletionLight := FALSE;
        (* MotorForward set on rising edge of firingComplete above *)

    ELSIF SensorWeight THEN
        (* ================================================================= *)
        (* STATION 3: WEIGHING                                                *)
        (* PUB006, PUB007, PUB008, PUB009                                     *)
        (* Motor stops; weightComplete triggers qualification check           *)
        (* ================================================================= *)
        state := ST_WEIGH;
        MotorForward := FALSE;
        CompletionLight := FALSE;

        (* Rising edge detection for weightComplete *)
        IF weightComplete AND NOT prevWeightComplete THEN
            prevWeightComplete := weightComplete;

            (* Qualification check: 100 <= weight <= 200 *)
            IF weight >= 100.0 AND weight <= 200.0 THEN
                (* Qualified: calculate firing temperature *)
                (* Linear interpolation: weight[100,200] -> temp[500,550] *)
                tmp_TempCalc := 500.0 + (weight - 100.0) * 0.5;
                firingTemp := tmp_TempCalc;
                kick := FALSE;
                MotorForward := TRUE;
            ELSE
                (* Unqualified: reject *)
                kick := TRUE;
                MotorForward := FALSE;
            END_IF;
        ELSE
            prevWeightComplete := weightComplete;
        END_IF;

    ELSIF SensorWash THEN
        (* ================================================================= *)
        (* STATION 2: CLEANING                                                *)
        (* PUB004, PUB005                                                     *)
        (* Motor stops; washComplete triggers forward                        *)
        (* ================================================================= *)
        state := ST_WASH;
        MotorForward := FALSE;
        CompletionLight := FALSE;
        kick := FALSE;  (* Reset kick on new product entering wash *)

    ELSIF SensorFeed THEN
        (* ================================================================= *)
        (* STATION 1: MATERIAL LOADING                                        *)
        (* PUB004                                                              *)
        (* SensorFeed detected → start motor forward                         *)
        (* ================================================================= *)
        state := ST_LOAD;
        MotorForward := TRUE;
        CompletionLight := FALSE;
        kick := FALSE;  (* Reset kick on new product *)

    ELSE
        (* No sensor active - product in transit or line empty *)
        (* Maintain current MotorForward state from completion signals *)
        (* MotorForward already set by rising edges above *)
        CompletionLight := FALSE;
    END_IF;

END_IF;

END_FUNCTION_BLOCK

(* ---- public-hard-06.raw_candidate_02.st ---- *)
(* ENGINEERING_CONTRACT
 * =============================================================================
 * Production Control - 5-Station Automated Line
 * =============================================================================
 * MODES:
 * - Manual (Mode=0): ForwardButton→MotorForward, ReverseButton→MotorReverse
 *   Interlock: MotorForward AND MotorReverse never simultaneous
 *   Activation: Button held; No retention; No explicit reset defined
 *
 * - Automatic (Mode=1): State-machine progression with sensor triggers
 *   States: LOAD→WASH→WEIGH→FIRE→OUTPUT (sequential forward flow)
 *
 * AUTOMATIC STATE TRANSITIONS:
 * - ST_LOAD: SensorFeed → MotorForward (retract, moves to next station)
 *   Reset: Automatic off, manual mode
 *
 * - ST_WASH: SensorWash → MotorStop
 *   Activation: washComplete → MotorForward
 *   Reset: Automatic off, manual mode
 *
 * - ST_WEIGH: SensorWeight → MotorStop
 *   Activation: weightComplete AND qualified(100≤weight≤200) → calc firingTemp, MotorForward
 *   Activation: weightComplete AND NOT qualified → kick latch ON
 *   Reset: Automatic off, manual mode; kick requires external reset (unspecified)
 *
 * - ST_FIRE: SensorFiring → MotorStop
 *   Activation: firingComplete → MotorForward
 *   Reset: Automatic off, manual mode
 *
 * - ST_OUTPUT: SensorOutput → MotorStop, CompletionLight:=SensorOutput
 *   Retention: CompletionLight held ON while SensorOutput=TRUE; OFF when FALSE
 *   Reset: Automatic off, manual mode (light follows sensor)
 *
 * FIRING TEMP CALCULATION:
 * - Linear: weight 100→200 maps to temp 500→550
 * - Formula: firingTemp = 500.0 + (weight - 100.0) * 0.5
 * - Only calculated once per qualified product (on weightComplete)
 * - Retained until next qualified product (unspecified reset)
 *
 * UNITS/BOUNDARIES:
 * - Weight: REAL, qualified range [100.0, 200.0] inclusive
 * - Temp: REAL, output range [500.0, 550.0] inclusive
 * - All sensors: BOOL, edge-triggered detection (sensor TRUE = product arrived)
 * =============================================================================
 *)

(* CONTRACT_RULES [{"kind":"hold_until_reset","output":"kick","set_input":"weightComplete","reset_input":null}] *)

TYPE StationState :
(
    ST_LOAD   := 0,
    ST_WASH   := 1,
    ST_WEIGH  := 2,
    ST_FIRE   := 3,
    ST_OUTPUT := 4
);
END_TYPE

FUNCTION_BLOCK ProductionControl
VAR_INPUT
    Mode            : BOOL;  (* 0=manual, 1=automatic *)
    ForwardButton   : BOOL;
    ReverseButton   : BOOL;
    SensorFeed      : BOOL;
    SensorWash      : BOOL;
    SensorWeight    : BOOL;
    SensorFiring    : BOOL;
    SensorOutput    : BOOL;
    washComplete    : BOOL;
    weightComplete  : BOOL;
    weight          : REAL;
    firingComplete  : BOOL;
END_VAR

VAR_OUTPUT
    MotorForward    : BOOL;
    MotorReverse    : BOOL;
    kick            : BOOL;
    CompletionLight : BOOL;
    firingTemp      : REAL;
END_VAR

VAR
    state               : StationState;
    prevWashComplete    : BOOL;
    prevWeightComplete  : BOOL;
    prevFiringComplete  : BOOL;
    tmp_Qualified       : BOOL;
    tmp_TempCalc        : REAL;
END_VAR

(* Initialize outputs to safe state *)
MotorForward    := FALSE;
MotorReverse    := FALSE;
kick            := kick;        (* Preserve retained state *)
CompletionLight := FALSE;
firingTemp      := firingTemp;  (* Preserve retained state *)

IF Mode = FALSE THEN
    (* ======================================================================= *)
    (* MANUAL MODE                                                             *)
    (* PUB001, PUB002, PUB003                                                  *)
    (* ======================================================================= *)
    (* Interlock: forward and reverse cannot be simultaneous *)
    IF ForwardButton AND NOT ReverseButton THEN
        MotorForward := TRUE;
        MotorReverse := FALSE;
    ELSIF ReverseButton AND NOT ForwardButton THEN
        MotorForward := FALSE;
        MotorReverse := TRUE;
    ELSE
        MotorForward := FALSE;
        MotorReverse := FALSE;
    END_IF;

    (* Reset state machine when entering manual mode *)
    state := ST_LOAD;

ELSIF Mode = TRUE THEN
    (* ======================================================================= *)
    (* AUTOMATIC MODE                                                          *)
    (* PUB004, PUB005, PUB006, PUB007, PUB008, PUB009, PUB010, PUB011, PUB012   *)
    (* ======================================================================= *)
    MotorReverse := FALSE;  (* Only forward in automatic mode *)

    (* Edge detection for completion signals *)
    IF washComplete AND NOT prevWashComplete THEN
        (* Rising edge on washComplete *)
        MotorForward := TRUE;
    END_IF;
    prevWashComplete := washComplete;

    IF firingComplete AND NOT prevFiringComplete THEN
        (* Rising edge on firingComplete *)
        MotorForward := TRUE;
    END_IF;
    prevFiringComplete := firingComplete;

    (* State machine based on current station detection *)
    IF SensorOutput THEN
        (* ================================================================= *)
        (* STATION 5: OUTPUT (Finished Product)                              *)
        (* PUB012                                                              *)
        (* Motor stops, CompletionLight follows sensor                       *)
        (* ================================================================= *)
        state := ST_OUTPUT;
        MotorForward := FALSE;
        CompletionLight := SensorOutput;  (* ON when product present *)

    ELSIF SensorFiring THEN
        (* ================================================================= *)
        (* STATION 4: FIRING                                                 *)
        (* PUB010, PUB011                                                     *)
        (* Motor stops; wait for firingComplete → forward                    *)
        (* ================================================================= *)
        state := ST_FIRE;
        MotorForward := FALSE;
        CompletionLight := FALSE;
        (* MotorForward set on rising edge of firingComplete above *)

    ELSIF SensorWeight THEN
        (* ================================================================= *)
        (* STATION 3: WEIGHING                                                *)
        (* PUB006, PUB007, PUB008, PUB009                                     *)
        (* Motor stops; weightComplete triggers qualification check           *)
        (* ================================================================= *)
        state := ST_WEIGH;
        MotorForward := FALSE;
        CompletionLight := FALSE;

        (* Rising edge detection for weightComplete *)
        IF weightComplete AND NOT prevWeightComplete THEN
            prevWeightComplete := weightComplete;

            (* Qualification check: 100 <= weight <= 200 *)
            IF weight >= 100.0 AND weight <= 200.0 THEN
                (* Qualified: calculate firing temperature *)
                (* Linear interpolation: weight[100,200] -> temp[500,550] *)
                tmp_TempCalc := 500.0 + (weight - 100.0) * 0.5;
                firingTemp := tmp_TempCalc;
                kick := FALSE;
                MotorForward := TRUE;
            ELSE
                (* Unqualified: reject *)
                kick := TRUE;
                MotorForward := FALSE;
            END_IF;
        ELSE
            prevWeightComplete := weightComplete;
        END_IF;

    ELSIF SensorWash THEN
        (* ================================================================= *)
        (* STATION 2: CLEANING                                                *)
        (* PUB004, PUB005                                                     *)
        (* Motor stops; washComplete triggers forward                        *)
        (* ================================================================= *)
        state := ST_WASH;
        MotorForward := FALSE;
        CompletionLight := FALSE;
        kick := FALSE;  (* Reset kick on new product entering wash *)

    ELSIF SensorFeed THEN
        (* ================================================================= *)
        (* STATION 1: MATERIAL LOADING                                        *)
        (* PUB004                                                              *)
        (* SensorFeed detected → start motor forward                         *)
        (* ================================================================= *)
        state := ST_LOAD;
        MotorForward := TRUE;
        CompletionLight := FALSE;
        kick := FALSE;  (* Reset kick on new product *)

    ELSE
        (* No sensor active - product in transit or line empty *)
        (* Maintain current MotorForward state from completion signals *)
        (* MotorForward already set by rising edges above *)
        CompletionLight := FALSE;
    END_IF;

END_IF;

END_FUNCTION_BLOCK

(* ---- public-hard-06.raw_candidate_03.st ---- *)
(* ENGINEERING_CONTRACT
 * =============================================================================
 * Production Control - 5-Station Automated Line
 * =============================================================================
 * MODES:
 * - Manual (Mode=0): ForwardButton→MotorForward, ReverseButton→MotorReverse
 *   Interlock: MotorForward AND MotorReverse never simultaneous
 *   Activation: Button held; No retention; No explicit reset defined
 *
 * - Automatic (Mode=1): State-machine progression with sensor triggers
 *   States: LOAD→WASH→WEIGH→FIRE→OUTPUT (sequential forward flow)
 *
 * AUTOMATIC STATE TRANSITIONS:
 * - ST_LOAD: SensorFeed → MotorForward (retract, moves to next station)
 *   Reset: Automatic off, manual mode
 *
 * - ST_WASH: SensorWash → MotorStop
 *   Activation: washComplete → MotorForward
 *   Reset: Automatic off, manual mode
 *
 * - ST_WEIGH: SensorWeight → MotorStop
 *   Activation: weightComplete AND qualified(100≤weight≤200) → calc firingTemp, MotorForward
 *   Activation: weightComplete AND NOT qualified → kick latch ON
 *   Reset: Automatic off, manual mode; kick requires external reset (unspecified)
 *
 * - ST_FIRE: SensorFiring → MotorStop
 *   Activation: firingComplete → MotorForward
 *   Reset: Automatic off, manual mode
 *
 * - ST_OUTPUT: SensorOutput → MotorStop, CompletionLight:=SensorOutput
 *   Retention: CompletionLight held ON while SensorOutput=TRUE; OFF when FALSE
 *   Reset: Automatic off, manual mode (light follows sensor)
 *
 * FIRING TEMP CALCULATION:
 * - Linear: weight 100→200 maps to temp 500→550
 * - Formula: firingTemp = 500.0 + (weight - 100.0) * 0.5
 * - Same-scan calculation when SensorWeight AND weightComplete both TRUE
 * - Retained until next qualified product (unspecified reset)
 *
 * UNITS/BOUNDARIES:
 * - Weight: REAL, qualified range [100.0, 200.0] inclusive
 * - Temp: REAL, output range [500.0, 550.0] inclusive
 * - All sensors: BOOL, level-triggered detection (sensor TRUE = product present)
 * =============================================================================
 *)

(* CONTRACT_RULES [] *)

TYPE StationState :
(
    ST_LOAD   := 0,
    ST_WASH   := 1,
    ST_WEIGH  := 2,
    ST_FIRE   := 3,
    ST_OUTPUT := 4
);
END_TYPE;

FUNCTION_BLOCK ProductionControl
VAR_INPUT
    Mode            : BOOL;  (* 0=manual, 1=automatic *)
    ForwardButton   : BOOL;
    ReverseButton   : BOOL;
    SensorFeed      : BOOL;
    SensorWash      : BOOL;
    SensorWeight    : BOOL;
    SensorFiring    : BOOL;
    SensorOutput    : BOOL;
    washComplete    : BOOL;
    weightComplete  : BOOL;
    weight          : REAL;
    firingComplete  : BOOL;
END_VAR

VAR_OUTPUT
    MotorForward    : BOOL;
    MotorReverse    : BOOL;
    kick             : BOOL;
    CompletionLight : BOOL;
    firingTemp      : REAL;
END_VAR

VAR
    state              : StationState;
    prevWashComplete   : BOOL;
    prevFiringComplete : BOOL;
END_VAR

(* Initialize outputs to safe state *)
MotorForward    := FALSE;
MotorReverse    := FALSE;
kick            := kick;        (* Preserve retained state *)
CompletionLight := FALSE;
firingTemp      := firingTemp;  (* Preserve retained state *)

IF Mode = FALSE THEN
    (* ======================================================================= *)
    (* MANUAL MODE                                                             *)
    (* PUB001, PUB002, PUB003                                                  *)
    (* ======================================================================= *)
    (* Interlock: forward and reverse cannot be simultaneous *)
    IF ForwardButton AND NOT ReverseButton THEN
        MotorForward := TRUE;
        MotorReverse := FALSE;
    ELSIF ReverseButton AND NOT ForwardButton THEN
        MotorForward := FALSE;
        MotorReverse := TRUE;
    ELSE
        MotorForward := FALSE;
        MotorReverse := FALSE;
    END_IF;

    (* Reset state machine when entering manual mode *)
    state := ST_LOAD;

ELSIF Mode = TRUE THEN
    (* ======================================================================= *)
    (* AUTOMATIC MODE                                                          *)
    (* PUB004, PUB005, PUB006, PUB007, PUB008, PUB009, PUB010, PUB011, PUB012   *)
    (* ======================================================================= *)
    MotorReverse := FALSE;  (* Only forward in automatic mode *)

    (* Edge detection for washComplete - rising edge triggers forward *)
    IF washComplete AND NOT prevWashComplete THEN
        MotorForward := TRUE;
    END_IF;
    prevWashComplete := washComplete;

    (* Edge detection for firingComplete - rising edge triggers forward *)
    IF firingComplete AND NOT prevFiringComplete THEN
        MotorForward := TRUE;
    END_IF;
    prevFiringComplete := firingComplete;

    (* State machine based on current station detection *)
    IF SensorOutput THEN
        (* ================================================================= *)
        (* STATION 5: OUTPUT (Finished Product)                              *)
        (* PUB012                                                              *)
        (* Motor stops, CompletionLight follows sensor                       *)
        (* ================================================================= *)
        state := ST_OUTPUT;
        MotorForward := FALSE;
        CompletionLight := SensorOutput;  (* ON when product present *)

    ELSIF SensorFiring THEN
        (* ================================================================= *)
        (* STATION 4: FIRING                                                 *)
        (* PUB010, PUB011                                                     *)
        (* Motor stops; wait for firingComplete → forward                    *)
        (* ================================================================= *)
        state := ST_FIRE;
        MotorForward := FALSE;
        CompletionLight := FALSE;
        (* MotorForward set on rising edge of firingComplete above *)

    ELSIF SensorWeight THEN
        (* ================================================================= *)
        (* STATION 3: WEIGHING                                                *)
        (* PUB006, PUB007, PUB008, PUB009                                     *)
        (* Motor stops; weightComplete triggers qualification check           *)
        (* ================================================================= *)
        state := ST_WEIGH;
        MotorForward := FALSE;
        CompletionLight := FALSE;

        (* Immediate calculation when weightComplete signal is received *)
        (* No edge delay - weightComplete is a one-shot from external process *)
        IF weightComplete THEN
            (* Qualification check: 100 <= weight <= 200 *)
            IF weight >= 100.0 AND weight <= 200.0 THEN
                (* Qualified: calculate firing temperature *)
                (* Linear interpolation: weight[100,200] -> temp[500,550] *)
                firingTemp := 500.0 + (weight - 100.0) * 0.5;
                kick := FALSE;
                MotorForward := TRUE;
            ELSE
                (* Unqualified: reject *)
                kick := TRUE;
                MotorForward := FALSE;
            END_IF;
        END_IF;

    ELSIF SensorWash THEN
        (* ================================================================= *)
        (* STATION 2: CLEANING                                                *)
        (* PUB004, PUB005                                                     *)
        (* Motor stops; washComplete triggers forward                        *)
        (* ================================================================= *)
        state := ST_WASH;
        MotorForward := FALSE;
        CompletionLight := FALSE;
        kick := FALSE;  (* Reset kick on new product entering wash *)

    ELSIF SensorFeed THEN
        (* ================================================================= *)
        (* STATION 1: MATERIAL LOADING                                        *)
        (* PUB004                                                              *)
        (* SensorFeed detected → start motor forward                         *)
        (* ================================================================= *)
        state := ST_LOAD;
        MotorForward := TRUE;
        CompletionLight := FALSE;
        kick := FALSE;  (* Reset kick on new product *)

    ELSE
        (* No sensor active - product in transit or line empty *)
        (* Maintain current MotorForward state from completion signals *)
        (* MotorForward already set by rising edges above *)
        CompletionLight := FALSE;
    END_IF;

END_IF;

END_FUNCTION_BLOCK

(* ---- public-hard-06.raw_candidate_04.st ---- *)
(* ENGINEERING_CONTRACT
 * Production Control - 5-Station Line
 * =============================================================================
 * MODES:
 * - Manual (Mode=0): ForwardButton→MotorForward, ReverseButton→MotorReverse
 *   Interlock: MotorForward AND MotorReverse never simultaneous
 *   Activation: Button held; No retention; No explicit reset defined
 *
 * - Automatic (Mode=1): State-machine progression with sensor triggers
 *   States: LOAD→WASH→WEIGH→FIRE→OUTPUT (sequential forward flow)
 *
 * AUTOMATIC STATE TRANSITIONS:
 * - ST_LOAD: SensorFeed → MotorForward (moves to cleaning station)
 * - ST_WASH: SensorWash → MotorStop; washComplete rising edge → MotorForward
 * - ST_WEIGH: SensorWeight → MotorStop; weightComplete rising edge:
 *   • weight in [100,200] → calc firingTemp (500+0.5*(w-100)), MotorForward
 *   • weight outside range → kick:=TRUE
 * - ST_FIRE: SensorFiring → MotorStop; firingComplete rising edge → MotorForward
 * - ST_OUTPUT: SensorOutput → MotorStop, CompletionLight:=SensorOutput
 *
 * UNITS/BOUNDARIES: Weight REAL in [100,200], Temp REAL in [500,550]
 * =============================================================================
 *)

(* CONTRACT_RULES [{"kind":"hold_until_reset","output":"kick","set_input":"weightComplete","reset_input":null}] *)

TYPE StationState :
(
    ST_LOAD   := 0,
    ST_WASH   := 1,
    ST_WEIGH  := 2,
    ST_FIRE   := 3,
    ST_OUTPUT := 4
);
END_TYPE;

FUNCTION_BLOCK ProductionControl
VAR_INPUT
    Mode            : BOOL;
    ForwardButton   : BOOL;
    ReverseButton   : BOOL;
    SensorFeed      : BOOL;
    SensorWash      : BOOL;
    SensorWeight    : BOOL;
    SensorFiring    : BOOL;
    SensorOutput    : BOOL;
    washComplete    : BOOL;
    weightComplete  : BOOL;
    weight          : REAL;
    firingComplete  : BOOL;
END_VAR

VAR_OUTPUT
    MotorForward    : BOOL;
    MotorReverse    : BOOL;
    kick            : BOOL;
    CompletionLight : BOOL;
    firingTemp      : REAL;
END_VAR

VAR
    state               : StationState;
    prevWashComplete    : BOOL;
    prevWeightComplete  : BOOL;
    prevFiringComplete  : BOOL;
    tmp_MotorForwardCmd : BOOL;
END_VAR

(* Rising edge detection - evaluate BEFORE any state transitions *)
VAR
    washCompleteRising   : BOOL;
    weightCompleteRising : BOOL;
    firingCompleteRising : BOOL;
END_VAR

washCompleteRising   := washComplete   AND NOT prevWashComplete;
weightCompleteRising := weightComplete AND NOT prevWeightComplete;
firingCompleteRising := firingComplete AND NOT prevFiringComplete;

(* Update previous states AFTER edge detection *)
prevWashComplete   := washComplete;
prevWeightComplete := weightComplete;
prevFiringComplete := firingComplete;

(* Default outputs - safety state *)
MotorForward    := FALSE;
MotorReverse    := FALSE;
CompletionLight := FALSE;

IF Mode = FALSE THEN
    (* ======================================================================= *)
    (* MANUAL MODE - PUB001, PUB002, PUB003                                    *)
    (* ======================================================================= *)
    IF ForwardButton AND NOT ReverseButton THEN
        MotorForward := TRUE;
        MotorReverse := FALSE;
    ELSIF ReverseButton AND NOT ForwardButton THEN
        MotorForward := FALSE;
        MotorReverse := TRUE;
    ELSE
        MotorForward := FALSE;
        MotorReverse := FALSE;
    END_IF;

    state := ST_LOAD;

ELSE
    (* ======================================================================= *)
    (* AUTOMATIC MODE - PUB004-PUB012                                           *)
    (* ======================================================================= *)
    MotorReverse := FALSE;

    (* Completion edges set motor forward command - takes priority *)
    IF washCompleteRising THEN
        tmp_MotorForwardCmd := TRUE;
    ELSIF firingCompleteRising THEN
        tmp_MotorForwardCmd := TRUE;
    ELSE
        tmp_MotorForwardCmd := FALSE;
    END_IF;

    (* Kick latch: activated on weightComplete rising edge per contract *)
    IF weightCompleteRising THEN
        IF weight >= 100.0 AND weight <= 200.0 THEN
            kick := FALSE;
        ELSE
            kick := TRUE;
        END_IF;
    END_IF;

    (* Firing temp: calculated on weightComplete rising edge for qualified weight *)
    IF weightCompleteRising THEN
        IF weight >= 100.0 AND weight <= 200.0 THEN
            firingTemp := 500.0 + (weight - 100.0) * 0.5;
        END_IF;
    END_IF;

    (* State machine based on sensor detection *)
    IF SensorOutput THEN
        state := ST_OUTPUT;
        tmp_MotorForwardCmd := FALSE;
        CompletionLight := TRUE;

    ELSIF SensorFiring THEN
        state := ST_FIRE;
        (* Only clear if no completion edge overrode *)
        IF NOT firingCompleteRising THEN
            tmp_MotorForwardCmd := FALSE;
        END_IF;
        CompletionLight := FALSE;

    ELSIF SensorWeight THEN
        state := ST_WEIGH;
        IF NOT weightCompleteRising THEN
            tmp_MotorForwardCmd := FALSE;
        END_IF;
        CompletionLight := FALSE;

    ELSIF SensorWash THEN
        state := ST_WASH;
        IF NOT washCompleteRising THEN
            tmp_MotorForwardCmd := FALSE;
        END_IF;
        CompletionLight := FALSE;

    ELSIF SensorFeed THEN
        state := ST_LOAD;
        tmp_MotorForwardCmd := TRUE;
        CompletionLight := FALSE;
        kick := FALSE;

    ELSE
        (* No sensor active - product in transit *)
        CompletionLight := FALSE;
    END_IF;

END_IF;

(* Apply accumulated motor forward command *)
MotorForward := tmp_MotorForwardCmd;

END_FUNCTION_BLOCK

(* ---- public-medium-01.candidate_01.st ---- *)
(* ENGINEERING_CONTRACT
 * PUB001: Mode selection - mode=FALSE selects Manual, mode=TRUE selects Automatic.
 * PUB002: Manual mode - read pumpGroup[].selection; write RunComd=TRUE on start for selected pumps.
 * PUB003: Automatic mode - sort 5 pumps by priority DESC, select top 3; write RunComd=TRUE for those pumps.
 * PUB004: Stop button - write RunComd=FALSE to all pumps regardless of mode (explicit reset).
 * Activation: R_TRIG on start/stop for single-scan edge detection (not level-triggered).
 * Retention: RunComd persists across scans until explicitly changed; no implicit state clear.
 * Priority rules: No specified simultaneous-operation conflict resolution; last command wins per scan.
 * Units: Priority is INT; no explicit range; 0 treated as lowest/skip. Lower array index wins ties.
 * Boundaries: Automatic mode selects exactly 3 pumps (or fewer if priority<=0); min 0 pumps selected.
 * CONTRACT_RULES [{"kind":"hold_until_reset","output":"pumpGroup","set_input":"start","reset_input":"stop"}]
 *)
FUNCTION_BLOCK FB_MultiPumpControl
VAR_INPUT
    mode  : BOOL;  // FALSE=Manual, TRUE=Automatic
    start : BOOL;
    stop  : BOOL;
END_VAR
VAR_IN_OUT
    pumpGroup : ARRAY[1..5] OF ST_Pump;
END_VAR
VAR
    startTrig  : R_TRIG;
    stopTrig   : R_TRIG;
END_VAR

// Rising-edge detection for start and stop buttons
startTrig(CLK := start);
stopTrig(CLK := stop);

// Stop button has highest priority - stops all pumps in any mode
IF stopTrig.Q THEN
    FOR 1 TO 5 DO
        pumpGroup[1].RunComd := FALSE;
        pumpGroup[2].RunComd := FALSE;
        pumpGroup[3].RunComd := FALSE;
        pumpGroup[4].RunComd := FALSE;
        pumpGroup[5].RunComd := FALSE;
    END_FOR;
    RETURN;
END_IF;

// Start command processed when stop is not active
IF startTrig.Q THEN
    IF mode = FALSE THEN
        // Manual mode: start selected pumps based on selection flag
        FOR 1 TO 5 DO
            pumpGroup[1].RunComd := pumpGroup[1].selection;
            pumpGroup[2].RunComd := pumpGroup[2].selection;
            pumpGroup[3].RunComd := pumpGroup[3].selection;
            pumpGroup[4].RunComd := pumpGroup[4].selection;
            pumpGroup[5].RunComd := pumpGroup[5].selection;
        END_FOR;
    ELSE
        // Automatic mode: select top 3 pumps by priority (highest priority first)
        VAR
            tmp_pumpCount   : INT := 0;
            tmp_priorities  : ARRAY[1..5] OF INT;
            tmp_indices     : ARRAY[1..5] OF INT;
            tmp_result      : ARRAY[1..3] OF INT;
            tmp_resultCount : INT := 0;
            i, j, tmp       : INT;
        END_VAR

        // Collect pumps with positive priority
        FOR i := 1 TO 5 DO
            IF pumpGroup[i].priority > 0 THEN
                tmp_pumpCount := tmp_pumpCount + 1;
                tmp_priorities[tmp_pumpCount] := pumpGroup[i].priority;
                tmp_indices[tmp_pumpCount] := i;
            END_IF;
        END_FOR;

        // Initialize result array
        FOR i := 1 TO 3 DO
            tmp_result[i] := 0;
        END_FOR;
        tmp_resultCount := 0;

        // Selection sort to find top 3 pumps by priority (descending)
        FOR i := 1 TO tmp_pumpCount DO
            VAR
                maxIdx : INT := i;
                maxVal : INT := tmp_priorities[i];
            END_VAR
            FOR j := i + 1 TO tmp_pumpCount DO
                IF tmp_priorities[j] > maxVal THEN
                    maxIdx  := j;
                    maxVal  := tmp_priorities[j];
                END_IF;
            END_FOR;
            // Swap to move max to position i
            tmp_priorities[maxIdx] := tmp_priorities[i];
            tmp_priorities[i]       := maxVal;
            tmp := tmp_indices[maxIdx];
            tmp_indices[maxIdx]     := tmp_indices[i];
            tmp_indices[i]          := tmp;

            // Record result (up to 3)
            IF tmp_resultCount < 3 THEN
                tmp_resultCount := tmp_resultCount + 1;
                tmp_result[tmp_resultCount] := tmp_indices[i];
            END_IF;
        END_FOR;

        // Apply run commands based on sorted selection
        FOR i := 1 TO 5 DO
            VAR
                isSelected : BOOL := FALSE;
            END_VAR
            FOR j := 1 TO tmp_resultCount DO
                IF tmp_result[j] = i THEN
                    isSelected := TRUE;
                    EXIT;
                END_IF;
            END_FOR;
            pumpGroup[i].RunComd := isSelected;
        END_FOR;
    END_IF;
END_IF;

END_FUNCTION_BLOCK

(* ---- public-medium-01.candidate_02.st ---- *)
(* ENGINEERING_CONTRACT
 * PUB001: Mode selection - mode=FALSE selects Manual, mode=TRUE selects Automatic.
 * PUB002: Manual mode - read pumpGroup[].selection; write RunComd=TRUE on start for selected pumps.
 * PUB003: Automatic mode - sort 5 pumps by priority DESC, select top 3; write RunComd=TRUE for those pumps.
 * PUB004: Stop button - write RunComd=FALSE to all pumps regardless of mode (explicit reset).
 * Activation: R_TRIG on start/stop for single-scan edge detection (not level-triggered).
 * Retention: RunComd persists across scans until explicitly changed; no implicit state clear.
 * Priority rules: No specified simultaneous-operation conflict resolution; last command wins per scan.
 * Units: Priority is INT; no explicit range; 0 or negative treated as skip. Lower array index wins ties.
 * Boundaries: Automatic mode selects up to 3 pumps with positive priority.
 * CONTRACT_RULES [{"kind":"hold_until_reset","output":"pumpGroup","set_input":"start","reset_input":"stop"}]
 *)
FUNCTION_BLOCK FB_MultiPumpControl
VAR_INPUT
    mode  : BOOL;  // FALSE=Manual, TRUE=Automatic
    start : BOOL;
    stop  : BOOL;
END_VAR
VAR_IN_OUT
    pumpGroup : ARRAY[1..5] OF ST_Pump;
END_VAR
VAR
    startTrig    : R_TRIG;
    stopTrig     : R_TRIG;
    tmp_pumpCount   : INT;
    tmp_priorities  : ARRAY[1..5] OF INT;
    tmp_indices     : ARRAY[1..5] OF INT;
    tmp_result      : ARRAY[1..3] OF INT;
    tmp_resultCount : INT;
    tmp_i, tmp_j, tmp_swap : INT;
    tmp_isSelected  : BOOL;
    tmp_maxIdx, tmp_maxVal : INT;
END_VAR

// Rising-edge detection for start and stop buttons
startTrig(CLK := start);
stopTrig(CLK := stop);

// Stop button has highest priority - stops all pumps in any mode
IF stopTrig.Q THEN
    FOR tmp_i := 1 TO 5 DO
        pumpGroup[tmp_i].RunComd := FALSE;
    END_FOR;
    RETURN;
END_IF;

// Start command processed when stop is not active
IF startTrig.Q THEN
    IF mode = FALSE THEN
        // Manual mode: start selected pumps based on selection flag
        FOR tmp_i := 1 TO 5 DO
            pumpGroup[tmp_i].RunComd := pumpGroup[tmp_i].selection;
        END_FOR;
    ELSE
        // Automatic mode: select top 3 pumps by priority (highest priority first)
        tmp_pumpCount := 0;

        // Collect pumps with positive priority
        FOR tmp_i := 1 TO 5 DO
            IF pumpGroup[tmp_i].priority > 0 THEN
                tmp_pumpCount := tmp_pumpCount + 1;
                tmp_priorities[tmp_pumpCount] := pumpGroup[tmp_i].priority;
                tmp_indices[tmp_pumpCount] := tmp_i;
            END_IF;
        END_FOR;

        // Initialize result array
        FOR tmp_i := 1 TO 3 DO
            tmp_result[tmp_i] := 0;
        END_FOR;
        tmp_resultCount := 0;

        // Selection sort to find top 3 pumps by priority (descending)
        FOR tmp_i := 1 TO tmp_pumpCount DO
            tmp_maxIdx := tmp_i;
            tmp_maxVal := tmp_priorities[tmp_i];
            FOR tmp_j := tmp_i + 1 TO tmp_pumpCount DO
                IF tmp_priorities[tmp_j] > tmp_maxVal THEN
                    tmp_maxIdx := tmp_j;
                    tmp_maxVal := tmp_priorities[tmp_j];
                END_IF;
            END_FOR;

            // Swap to move max to position tmp_i
            tmp_priorities[tmp_maxIdx] := tmp_priorities[tmp_i];
            tmp_priorities[tmp_i] := tmp_maxVal;
            tmp_swap := tmp_indices[tmp_maxIdx];
            tmp_indices[tmp_maxIdx] := tmp_indices[tmp_i];
            tmp_indices[tmp_i] := tmp_swap;

            // Record result (up to 3)
            IF tmp_resultCount < 3 THEN
                tmp_resultCount := tmp_resultCount + 1;
                tmp_result[tmp_resultCount] := tmp_indices[tmp_i];
            END_IF;
        END_FOR;

        // Apply run commands based on sorted selection
        FOR tmp_i := 1 TO 5 DO
            tmp_isSelected := FALSE;
            FOR tmp_j := 1 TO tmp_resultCount DO
                IF tmp_result[tmp_j] = tmp_i THEN
                    tmp_isSelected := TRUE;
                    EXIT;
                END_IF;
            END_FOR;
            pumpGroup[tmp_i].RunComd := tmp_isSelected;
        END_FOR;
    END_IF;
END_IF;

END_FUNCTION_BLOCK
